TYPE ST_EL3356CoeReadData :
STRUCT
	wIdx: WORD;
	bySubIdx: BYTE;
	bReadOK: BOOL;
	dwData: DWORD;
	nSize: UDINT;
END_STRUCT
END_TYPE

(* stored: Version 1.1.0.1, ProductVersion 3.1.4024.15
   DUT ST_EL3356CoeReadData: Id {6f13aab1-4fea-4de0-8a26-7025aa170177} *)
